(* Schneider Machine Expert - Basic project mojokerto-rev7, file version 2.9.0.0 *)
(* ProjectInformations: Name=New project *)

HARDWARE
  Cpu 0: TM221CE24R
  EthernetConfiguration: NetworkName=M221, IpAllocationMode=FixedAddress, IpAddress=192.168.1.113, SubnetMask=255.255.255.0
  SerialLineConfiguration: Baud=Baud19200, Parity=ParityNone, DataBits=DataBits8, StopBits=StopBits1, PhysicalMedium=PhysicalMediumRs485, TransmissionMode=TransmissionModeIoScannerRtu
  MastTask: UsePeriodScanMode=false, PeriodScan=100
  FastTask: Period=255
  CpuBehavior: StartingMode=StartAsPreviousState, AutoSaveRamOnEeprom=true, WatchdogPeriod=250

SYMBOLS  (address, symbol, comment, settings)
  %M10      VSD1_START  "VSD1 START dari FUXA (pulse)"
  %M11      VSD1_STOP  "VSD1 STOP dari FUXA (pulse)"
  %M12      VSD2_START  "VSD2 START dari FUXA (pulse)"
  %M13      VSD2_STOP  "VSD2 STOP dari FUXA (pulse)"
  %M14      VSD3_START  "VSD3 START dari FUXA (pulse)"
  %M15      VSD3_STOP  "VSD3 STOP dari FUXA (pulse)"
  %M16      VSD4_START  "VSD4 START dari FUXA (pulse)"
  %M17      VSD4_STOP  "VSD4 STOP dari FUXA (pulse)"
  %M18      VSD5_START  "VSD5 START dari FUXA (pulse)"
  %M19      VSD5_STOP  "VSD5 STOP dari FUXA (pulse)"
  %M20      VSD1_RUN_CMD  "VSD1 output RUN aktif"
  %M21      VSD2_RUN_CMD  "VSD2 output RUN aktif"
  %M22      VSD3_RUN_CMD  "VSD3 output RUN aktif"
  %M23      VSD4_RUN_CMD  "VSD4 output RUN aktif"
  %M24      VSD5_RUN_CMD  "VSD5 output RUN aktif"
  %M25      VSD1_RUNNING  "VSD1 berjalan (SW b2)"
  %M26      VSD2_RUNNING  "VSD2 berjalan (SW b2)"
  %M27      VSD3_RUNNING  "VSD3 berjalan (SW b2)"
  %M28      VSD4_RUNNING  "VSD4 berjalan (SW b2)"
  %M29      VSD5_RUNNING  "VSD5 berjalan (SW b2)"
  %M30      MODE_REMOTE  "1 = selector REMOTE (SCADA), 0 = LOCAL (PB panel)"
  %M31      MODE_ESTOP_OK  "Salinan %I0.1 untuk FUXA: 1 = e-stop sehat"
  %M40      VSD1_FAULT  "VSD1 fault (SW b3, comm OK)"
  %M41      VSD2_FAULT  "VSD2 fault (SW b3, comm OK)"
  %M42      VSD3_FAULT  "VSD3 fault (SW b3, comm OK)"
  %M43      VSD4_FAULT  "VSD4 fault (SW b3, comm OK)"
  %M44      VSD5_FAULT  "VSD5 fault (SW b3, comm OK)"
  %M45      VSD1_WARN  "VSD1 warning (SW b7)"
  %M46      VSD2_WARN  "VSD2 warning (SW b7)"
  %M47      VSD3_WARN  "VSD3 warning (SW b7)"
  %M48      VSD4_WARN  "VSD4 warning (SW b7)"
  %M49      VSD5_WARN  "VSD5 warning (SW b7)"
  %M50      VSD1_REMOTE  "VSD1 di REMOTE (SW b9)"
  %M51      VSD2_REMOTE  "VSD2 di REMOTE (SW b9)"
  %M52      VSD3_REMOTE  "VSD3 di REMOTE (SW b9)"
  %M53      VSD4_REMOTE  "VSD4 di REMOTE (SW b9)"
  %M54      VSD5_REMOTE  "VSD5 di REMOTE (SW b9)"
  %M60      VSD1_COMM_OK  "VSD1 IOScanner status = 2"
  %M61      VSD2_COMM_OK  "VSD2 IOScanner status = 2"
  %M62      VSD3_COMM_OK  "VSD3 IOScanner status = 2"
  %M63      VSD4_COMM_OK  "VSD4 IOScanner status = 2"
  %M64      VSD5_COMM_OK  "VSD5 IOScanner status = 2"
  %M65      FLOW_COMM_OK  "Flow meter IOScanner status = 2"
  %M70      VSD1_COMM_LOST  "VSD1 alarm komunikasi putus"
  %M71      VSD2_COMM_LOST  "VSD2 alarm komunikasi putus"
  %M72      VSD3_COMM_LOST  "VSD3 alarm komunikasi putus"
  %M73      VSD4_COMM_LOST  "VSD4 alarm komunikasi putus"
  %M74      VSD5_COMM_LOST  "VSD5 alarm komunikasi putus"
  %M75      FLOW_COMM_LOST  "Flow meter alarm komunikasi putus"
  %M80      FLOW_PIPE_EMPTY  "Flow: pipa kosong"
  %M81      FLOW_COIL_ERR  "Flow: coils excitation error"
  %M82      FLOW_MIN  "Flow: di bawah MIN"
  %M83      FLOW_MAX  "Flow: di atas MAX"
  %M90      VSD3_INSTALLED  "1 = VSD3 sudah terpasang, alarm comm lost VSD3 aktif"
  %M99      WORD_SWAP  "0 = tukar word 32-bit (default), 1 = lurus"
  %M111     RETRY_PULSE  "Pulse auto-retry IOScanner (rev5)"
  %M112     S6_PREV  "%S6 scan sebelumnya (deteksi sisi naik)"
  %S6       SB_TB1S  "Time base of 1 s generated by an internal clock"
  %S13      SB_FIRSTRUN  "Indicates the first controller cycle in RUN mode"
  %S110     SB_IOSCAN1RESET  "Set to 1 to reset the IOScanner on Serial Line 1"
  %SW210    SW_IOSCAN1STATUS  "Contains the IOScanner status of Serial Line 1"
  %MW990    SP_MIN  "Setpoint minimum Hz x10"
  %MW991    SP_MAX  "Setpoint maksimum Hz x10"
  %MW1000   VSD1_SW  "VSD1 status word"
  %MW1001   VSD1_FREQ  "VSD1 frekuensi Hz x10"
  %MW1002   VSD1_CURRENT  "VSD1 arus A x10"
  %MW1003   VSD1_DCBUS  "VSD1 DC bus V"
  %MW1004   VSD1_VOUT  "VSD1 Vout V"
  %MW1005   VSD1_REF_RB  "VSD1 ref1 terbaca Hz x10"
  %MW1006   VSD1_SP  "VSD1 setpoint dari FUXA Hz x10"
  %MW1020   VSD2_SW  "VSD2 status word"
  %MW1021   VSD2_FREQ  "VSD2 frekuensi Hz x10"
  %MW1022   VSD2_CURRENT  "VSD2 arus A x10"
  %MW1023   VSD2_DCBUS  "VSD2 DC bus V"
  %MW1024   VSD2_VOUT  "VSD2 Vout V"
  %MW1025   VSD2_REF_RB  "VSD2 ref1 terbaca Hz x10"
  %MW1026   VSD2_SP  "VSD2 setpoint dari FUXA Hz x10"
  %MW1040   VSD3_SW  "VSD3 status word"
  %MW1041   VSD3_FREQ  "VSD3 frekuensi Hz x10"
  %MW1042   VSD3_CURRENT  "VSD3 arus A x10"
  %MW1043   VSD3_DCBUS  "VSD3 DC bus V"
  %MW1044   VSD3_VOUT  "VSD3 Vout V"
  %MW1045   VSD3_REF_RB  "VSD3 ref1 terbaca Hz x10"
  %MW1046   VSD3_SP  "VSD3 setpoint dari FUXA Hz x10"
  %MW1060   VSD4_SW  "VSD4 status word"
  %MW1061   VSD4_FREQ  "VSD4 frekuensi Hz x10"
  %MW1062   VSD4_CURRENT  "VSD4 arus A x10"
  %MW1063   VSD4_DCBUS  "VSD4 DC bus V"
  %MW1064   VSD4_VOUT  "VSD4 Vout V"
  %MW1065   VSD4_REF_RB  "VSD4 ref1 terbaca Hz x10"
  %MW1066   VSD4_SP  "VSD4 setpoint dari FUXA Hz x10"
  %MW1080   VSD5_SW  "VSD5 status word"
  %MW1081   VSD5_FREQ  "VSD5 frekuensi Hz x10"
  %MW1082   VSD5_CURRENT  "VSD5 arus A x10"
  %MW1083   VSD5_DCBUS  "VSD5 DC bus V"
  %MW1084   VSD5_VOUT  "VSD5 Vout V"
  %MW1085   VSD5_REF_RB  "VSD5 ref1 terbaca Hz x10"
  %MW1086   VSD5_SP  "VSD5 setpoint dari FUXA Hz x10"
  %MW1112   FLOW_TP_INFO  "T+ MSB overflow LSB desimal"
  %MW1113   FLOW_TN_INFO  "T- info"
  %MW1114   FLOW_FLAGS12  "Flag 1/2 reg 0020"
  %MW1115   FLOW_ALARMS  "Jumlah alarm"
  %MW1116   FLOW_BATT  "Baterai %"
  %MW1117   FLOW_FLAGS34  "Flag 3/4 reg 0051"
  %MW1600   VSD1_IOS_STAT  "VSD1 status device IOScanner"
  %MW1601   VSD2_IOS_STAT  "VSD2 status device IOScanner"
  %MW1602   VSD3_IOS_STAT  "VSD3 status device IOScanner"
  %MW1603   FLOW_IOS_STAT  "Flow status device IOScanner"
  %MW1604   VSD4_IOS_STAT  "VSD4 status device IOScanner"
  %MW1605   VSD5_IOS_STAT  "VSD5 status device IOScanner"
  %MW1606   IOS_SL1_STATE  "%SW210: 0 stop 1 init 2 OK 3 sebagian 4 suspend"
  %MW1610   RETRY_SEC_CNT  "Hitungan detik auto-retry IOScanner"
  %MW1611   IOS_RESET_COUNT  "Jumlah reset IOScanner SL1 oleh program"
  %I0.0     SEL_REMOTE  "Selector panel: 1 = REMOTE (start/stop SCADA), 0 = LOCAL (PB panel)"
  %I0.1     ESTOP_OK  "E-stop, kontak NC: 1 = sehat"
  %I0.2     VSD1_PB_ON  "PB ON VSD1 di panel (NO), aktif di LOCAL"
  %I0.3     VSD1_PB_OFF  "PB OFF VSD1 di panel (NC), aktif di LOCAL dan REMOTE, 0 = stop"
  %I0.4     VSD2_PB_ON  "PB ON VSD2 di panel (NO), aktif di LOCAL"
  %I0.5     VSD2_PB_OFF  "PB OFF VSD2 di panel (NC), aktif di LOCAL dan REMOTE, 0 = stop"
  %I0.6     VSD3_PB_ON  "PB ON VSD3 di panel (NO), aktif di LOCAL"
  %I0.7     VSD3_PB_OFF  "PB OFF VSD3 di panel (NC), aktif di LOCAL dan REMOTE, 0 = stop"
  %I0.8     VSD4_PB_ON  "PB ON VSD4 di panel (NO), aktif di LOCAL"
  %I0.9     VSD4_PB_OFF  "PB OFF VSD4 di panel (NC), aktif di LOCAL dan REMOTE, 0 = stop"
  %I0.10    VSD5_PB_ON  "PB ON VSD5 di panel (NO), aktif di LOCAL"
  %I0.11    VSD5_PB_OFF  "PB OFF VSD5 di panel (NC), aktif di LOCAL dan REMOTE, 0 = stop"
  %Q0.0     VSD1_RUN  "Ke DI start VSD1 (ACS550), hardwired"
  %Q0.1     VSD2_RUN  "Ke DI start VSD2 (ACS580), hardwired"
  %Q0.2     VSD3_RUN  "Ke DI start VSD3 (ACS580), hardwired"
  %Q0.3     VSD4_RUN  "Ke DI start VSD4 (ACS580), hardwired"
  %Q0.4     VSD5_RUN  "Ke DI start VSD5 (ACS580), hardwired"
  %IWN100.0.0   [Channel=SW_REF_ACT]
  %IWN100.0.1   [Channel=SW_REF_ACT]
  %IWN100.0.2   [Channel=SW_REF_ACT]
  %IWN100.0.3   [Channel=SW_REF_ACT]
  %IWN100.1.0   [Channel=PAR_0103_0111]
  %IWN100.1.1   [Channel=PAR_0103_0111]
  %IWN100.1.2   [Channel=PAR_0103_0111]
  %IWN100.1.3   [Channel=PAR_0103_0111]
  %IWN100.1.4   [Channel=PAR_0103_0111]
  %IWN100.1.5   [Channel=PAR_0103_0111]
  %IWN100.1.6   [Channel=PAR_0103_0111]
  %IWN100.1.7   [Channel=PAR_0103_0111]
  %IWN100.1.8   [Channel=PAR_0103_0111]
  %IWN101.0.0   [Channel=SW_REF_ACT]
  %IWN101.0.1   [Channel=SW_REF_ACT]
  %IWN101.0.2   [Channel=SW_REF_ACT]
  %IWN101.0.3   [Channel=SW_REF_ACT]
  %IWN101.1.0   [Channel=CURRENT_32]
  %IWN101.1.1   [Channel=CURRENT_32]
  %IWN101.2.0   [Channel=DC_BUS]
  %IWN101.3.0   [Channel=VOUT]
  %IWN102.0.0   [Channel=SW_REF_ACT]
  %IWN102.0.1   [Channel=SW_REF_ACT]
  %IWN102.0.2   [Channel=SW_REF_ACT]
  %IWN102.0.3   [Channel=SW_REF_ACT]
  %IWN102.1.0   [Channel=CURRENT_32]
  %IWN102.1.1   [Channel=CURRENT_32]
  %IWN102.2.0   [Channel=DC_BUS]
  %IWN102.3.0   [Channel=VOUT]
  %IWN103.0.0   [Channel=FLOW_TOT_FLAGS]
  %IWN103.0.1   [Channel=FLOW_TOT_FLAGS]
  %IWN103.0.2   [Channel=FLOW_TOT_FLAGS]
  %IWN103.0.3   [Channel=FLOW_TOT_FLAGS]
  %IWN103.0.4   [Channel=FLOW_TOT_FLAGS]
  %IWN103.0.5   [Channel=FLOW_TOT_FLAGS]
  %IWN103.0.6   [Channel=FLOW_TOT_FLAGS]
  %IWN103.0.7   [Channel=FLOW_TOT_FLAGS]
  %IWN103.0.8   [Channel=FLOW_TOT_FLAGS]
  %IWN103.0.9   [Channel=FLOW_TOT_FLAGS]
  %IWN103.0.10   [Channel=FLOW_TOT_FLAGS]
  %IWN103.0.11   [Channel=FLOW_TOT_FLAGS]
  %IWN103.0.12   [Channel=FLOW_TOT_FLAGS]
  %IWN103.0.13   [Channel=FLOW_TOT_FLAGS]
  %IWN103.0.14   [Channel=FLOW_TOT_FLAGS]
  %IWN103.0.15   [Channel=FLOW_TOT_FLAGS]
  %IWN103.0.16   [Channel=FLOW_TOT_FLAGS]
  %IWN103.0.17   [Channel=FLOW_TOT_FLAGS]
  %IWN103.0.18   [Channel=FLOW_TOT_FLAGS]
  %IWN103.1.0   [Channel=BATT_ALM_LPS]
  %IWN103.1.1   [Channel=BATT_ALM_LPS]
  %IWN103.1.2   [Channel=BATT_ALM_LPS]
  %IWN103.1.3   [Channel=BATT_ALM_LPS]
  %IWN103.1.4   [Channel=BATT_ALM_LPS]
  %IWN103.1.5   [Channel=BATT_ALM_LPS]
  %IWN103.1.6   [Channel=BATT_ALM_LPS]
  %IWN103.1.7   [Channel=BATT_ALM_LPS]
  %IWN103.1.8   [Channel=BATT_ALM_LPS]
  %IWN103.1.9   [Channel=BATT_ALM_LPS]
  %IWN103.2.0   [Channel=FLAGS_3_4]
  %IWN104.0.0   [Channel=SW_REF_ACT]
  %IWN104.0.1   [Channel=SW_REF_ACT]
  %IWN104.0.2   [Channel=SW_REF_ACT]
  %IWN104.0.3   [Channel=SW_REF_ACT]
  %IWN104.1.0   [Channel=CURRENT_32]
  %IWN104.1.1   [Channel=CURRENT_32]
  %IWN104.2.0   [Channel=DC_BUS]
  %IWN104.3.0   [Channel=VOUT]
  %IWN105.0.0   [Channel=SW_REF_ACT]
  %IWN105.0.1   [Channel=SW_REF_ACT]
  %IWN105.0.2   [Channel=SW_REF_ACT]
  %IWN105.0.3   [Channel=SW_REF_ACT]
  %IWN105.1.0   [Channel=CURRENT_32]
  %IWN105.1.1   [Channel=CURRENT_32]
  %IWN105.2.0   [Channel=DC_BUS]
  %IWN105.3.0   [Channel=VOUT]
  %QWN100.2.0   [Channel=REF1_WRITE]
  %QWN101.4.0   [Channel=REF1_WRITE]
  %QWN102.4.0   [Channel=REF1_WRITE]
  %QWN104.4.0   [Channel=REF1_WRITE]
  %QWN105.4.0   [Channel=REF1_WRITE]

POU Mojokerto
  (* SectionNumber=0 *)

// Rung 0: INIT
// Cold start: batas setpoint default 0..50,0 Hz (x10)
  LD %S13                 (* SB_FIRSTRUN - Siklus pertama setelah start *)
  [ %MW990 := 0 ]         (* SP_MIN - SP_MIN Hz x10 *)
  [ %MW991 := 500 ]       (* SP_MAX - SP_MAX Hz x10 *)
  // as ST:
  //   IF SB_FIRSTRUN THEN SP_MIN := 0; END_IF;
  //   IF SB_FIRSTRUN THEN SP_MAX := 500; END_IF;

// Rung 1: RAW_VSD1
// Salin data IOScanner VSD1 (ACS550, slave ID 1) ke %MW1300
  LD 1                    (* Selalu *)
  [ %MW1300 := %IWN100.0.0 ](* ref1 *)
  [ %MW1301 := %IWN100.0.1 ](* ref2 *)
  [ %MW1302 := %IWN100.0.2 ](* status word *)
  [ %MW1303 := %IWN100.0.3 ](* act1 *)
  [ %MW1304 := %IWN100.1.0 ](* par 0103 *)
  [ %MW1305 := %IWN100.1.1 ](* par 0104 *)
  [ %MW1306 := %IWN100.1.2 ](* par 0105 *)
  [ %MW1307 := %IWN100.1.3 ](* par 0106 *)
  [ %MW1308 := %IWN100.1.4 ](* par 0107 *)
  [ %MW1309 := %IWN100.1.5 ](* par 0108 *)
  [ %MW1310 := %IWN100.1.6 ](* par 0109 *)
  [ %MW1311 := %IWN100.1.7 ](* par 0110 *)
  [ %MW1312 := %IWN100.1.8 ](* par 0111 *)
  [ %MW1600 := %IWNS100 ] (* VSD1_IOS_STAT - status device IOScanner (2 = OK) *)
  // as ST:
  //   %MW1300 := %IWN100.0.0;
  //   %MW1301 := %IWN100.0.1;
  //   %MW1302 := %IWN100.0.2;
  //   %MW1303 := %IWN100.0.3;
  //   %MW1304 := %IWN100.1.0;
  //   %MW1305 := %IWN100.1.1;
  //   %MW1306 := %IWN100.1.2;
  //   %MW1307 := %IWN100.1.3;
  //   %MW1308 := %IWN100.1.4;
  //   %MW1309 := %IWN100.1.5;
  //   %MW1310 := %IWN100.1.6;
  //   %MW1311 := %IWN100.1.7;
  //   %MW1312 := %IWN100.1.8;
  //   VSD1_IOS_STAT := %IWNS100;

// Rung 2: RAW_VSD2
// Salin data IOScanner VSD2 (ACS580, slave ID 2) ke %MW1340
  LD 1                    (* Selalu *)
  [ %MW1340 := %IWN101.0.0 ](* ref1 *)
  [ %MW1341 := %IWN101.0.1 ](* ref2 *)
  [ %MW1342 := %IWN101.0.2 ](* status word *)
  [ %MW1343 := %IWN101.0.3 ](* act1 *)
  [ %MW1344 := %IWN101.1.0 ](* 01.07 arus word 1 *)
  [ %MW1345 := %IWN101.1.1 ](* 01.07 arus word 2 *)
  [ %MW1346 := %IWN101.2.0 ](* 01.11 DC bus *)
  [ %MW1347 := %IWN101.3.0 ](* 01.13 Vout *)
  [ %MW1601 := %IWNS101 ] (* VSD2_IOS_STAT - status device IOScanner (2 = OK) *)
  // as ST:
  //   %MW1340 := %IWN101.0.0;
  //   %MW1341 := %IWN101.0.1;
  //   %MW1342 := %IWN101.0.2;
  //   %MW1343 := %IWN101.0.3;
  //   %MW1344 := %IWN101.1.0;
  //   %MW1345 := %IWN101.1.1;
  //   %MW1346 := %IWN101.2.0;
  //   %MW1347 := %IWN101.3.0;
  //   VSD2_IOS_STAT := %IWNS101;

// Rung 3: RAW_VSD3
// Salin data IOScanner VSD3 (ACS580, slave ID 3) ke %MW1380
  LD 1                    (* Selalu *)
  [ %MW1380 := %IWN102.0.0 ](* ref1 *)
  [ %MW1381 := %IWN102.0.1 ](* ref2 *)
  [ %MW1382 := %IWN102.0.2 ](* status word *)
  [ %MW1383 := %IWN102.0.3 ](* act1 *)
  [ %MW1384 := %IWN102.1.0 ](* 01.07 arus word 1 *)
  [ %MW1385 := %IWN102.1.1 ](* 01.07 arus word 2 *)
  [ %MW1386 := %IWN102.2.0 ](* 01.11 DC bus *)
  [ %MW1387 := %IWN102.3.0 ](* 01.13 Vout *)
  [ %MW1602 := %IWNS102 ] (* VSD3_IOS_STAT - status device IOScanner (2 = OK) *)
  // as ST:
  //   %MW1380 := %IWN102.0.0;
  //   %MW1381 := %IWN102.0.1;
  //   %MW1382 := %IWN102.0.2;
  //   %MW1383 := %IWN102.0.3;
  //   %MW1384 := %IWN102.1.0;
  //   %MW1385 := %IWN102.1.1;
  //   %MW1386 := %IWN102.2.0;
  //   %MW1387 := %IWN102.3.0;
  //   VSD3_IOS_STAT := %IWNS102;

// Rung 4: RAW_VSD4
// Salin data IOScanner VSD4 (ACS580, slave ID 5) ke %MW1460
  LD 1                    (* Selalu *)
  [ %MW1460 := %IWN104.0.0 ](* ref1 *)
  [ %MW1461 := %IWN104.0.1 ](* ref2 *)
  [ %MW1462 := %IWN104.0.2 ](* status word *)
  [ %MW1463 := %IWN104.0.3 ](* act1 *)
  [ %MW1464 := %IWN104.1.0 ](* 01.07 arus word 1 *)
  [ %MW1465 := %IWN104.1.1 ](* 01.07 arus word 2 *)
  [ %MW1466 := %IWN104.2.0 ](* 01.11 DC bus *)
  [ %MW1467 := %IWN104.3.0 ](* 01.13 Vout *)
  [ %MW1604 := %IWNS104 ] (* VSD4_IOS_STAT - status device IOScanner (2 = OK) *)
  // as ST:
  //   %MW1460 := %IWN104.0.0;
  //   %MW1461 := %IWN104.0.1;
  //   %MW1462 := %IWN104.0.2;
  //   %MW1463 := %IWN104.0.3;
  //   %MW1464 := %IWN104.1.0;
  //   %MW1465 := %IWN104.1.1;
  //   %MW1466 := %IWN104.2.0;
  //   %MW1467 := %IWN104.3.0;
  //   VSD4_IOS_STAT := %IWNS104;

// Rung 5: RAW_VSD5
// Salin data IOScanner VSD5 (ACS580, slave ID 6) ke %MW1500
  LD 1                    (* Selalu *)
  [ %MW1500 := %IWN105.0.0 ](* ref1 *)
  [ %MW1501 := %IWN105.0.1 ](* ref2 *)
  [ %MW1502 := %IWN105.0.2 ](* status word *)
  [ %MW1503 := %IWN105.0.3 ](* act1 *)
  [ %MW1504 := %IWN105.1.0 ](* 01.07 arus word 1 *)
  [ %MW1505 := %IWN105.1.1 ](* 01.07 arus word 2 *)
  [ %MW1506 := %IWN105.2.0 ](* 01.11 DC bus *)
  [ %MW1507 := %IWN105.3.0 ](* 01.13 Vout *)
  [ %MW1605 := %IWNS105 ] (* VSD5_IOS_STAT - status device IOScanner (2 = OK) *)
  // as ST:
  //   %MW1500 := %IWN105.0.0;
  //   %MW1501 := %IWN105.0.1;
  //   %MW1502 := %IWN105.0.2;
  //   %MW1503 := %IWN105.0.3;
  //   %MW1504 := %IWN105.1.0;
  //   %MW1505 := %IWN105.1.1;
  //   %MW1506 := %IWN105.2.0;
  //   %MW1507 := %IWN105.3.0;
  //   VSD5_IOS_STAT := %IWNS105;

// Rung 6: RAW_FLOW
// Salin data IOScanner flow meter MV145 (slave ID 4) ke %MW1420
  LD 1                    (* Selalu *)
  [ %MW1420 := %IWN103.0.0 ](* MV145 reg 0002 *)
  [ %MW1421 := %IWN103.0.1 ](* MV145 reg 0003 *)
  [ %MW1422 := %IWN103.0.2 ](* MV145 reg 0004 *)
  [ %MW1423 := %IWN103.0.3 ](* MV145 reg 0005 *)
  [ %MW1424 := %IWN103.0.4 ](* MV145 reg 0006 *)
  [ %MW1425 := %IWN103.0.5 ](* MV145 reg 0007 *)
  [ %MW1426 := %IWN103.0.6 ](* MV145 reg 0008 *)
  [ %MW1427 := %IWN103.0.7 ](* MV145 reg 0009 *)
  [ %MW1428 := %IWN103.0.8 ](* MV145 reg 0010 *)
  [ %MW1429 := %IWN103.0.9 ](* MV145 reg 0011 *)
  [ %MW1430 := %IWN103.0.10 ](* MV145 reg 0012 *)
  [ %MW1431 := %IWN103.0.11 ](* MV145 reg 0013 *)
  [ %MW1432 := %IWN103.0.12 ](* MV145 reg 0014 *)
  [ %MW1433 := %IWN103.0.13 ](* MV145 reg 0015 *)
  [ %MW1434 := %IWN103.0.14 ](* MV145 reg 0016 *)
  [ %MW1435 := %IWN103.0.15 ](* MV145 reg 0017 *)
  [ %MW1436 := %IWN103.0.16 ](* MV145 reg 0018 *)
  [ %MW1437 := %IWN103.0.17 ](* MV145 reg 0019 *)
  [ %MW1438 := %IWN103.0.18 ](* MV145 reg 0020 *)
  [ %MW1440 := %IWN103.1.0 ](* MV145 reg 0027 *)
  [ %MW1441 := %IWN103.1.1 ](* MV145 reg 0028 *)
  [ %MW1442 := %IWN103.1.2 ](* MV145 reg 0029 *)
  [ %MW1443 := %IWN103.1.3 ](* MV145 reg 0030 *)
  [ %MW1444 := %IWN103.1.4 ](* MV145 reg 0031 *)
  [ %MW1445 := %IWN103.1.5 ](* MV145 reg 0032 *)
  [ %MW1446 := %IWN103.1.6 ](* MV145 reg 0033 *)
  [ %MW1447 := %IWN103.1.7 ](* MV145 reg 0034 *)
  [ %MW1448 := %IWN103.1.8 ](* MV145 reg 0035 *)
  [ %MW1449 := %IWN103.1.9 ](* MV145 reg 0036 *)
  [ %MW1450 := %IWN103.2.0 ](* MV145 reg 0051 *)
  [ %MW1603 := %IWNS103 ] (* FLOW_IOS_STAT - status device IOScanner flow (2 = OK) *)
  // as ST:
  //   %MW1420 := %IWN103.0.0;
  //   %MW1421 := %IWN103.0.1;
  //   %MW1422 := %IWN103.0.2;
  //   %MW1423 := %IWN103.0.3;
  //   %MW1424 := %IWN103.0.4;
  //   %MW1425 := %IWN103.0.5;
  //   %MW1426 := %IWN103.0.6;
  //   %MW1427 := %IWN103.0.7;
  //   %MW1428 := %IWN103.0.8;
  //   %MW1429 := %IWN103.0.9;
  //   %MW1430 := %IWN103.0.10;
  //   %MW1431 := %IWN103.0.11;
  //   %MW1432 := %IWN103.0.12;
  //   %MW1433 := %IWN103.0.13;
  //   %MW1434 := %IWN103.0.14;
  //   %MW1435 := %IWN103.0.15;
  //   %MW1436 := %IWN103.0.16;
  //   %MW1437 := %IWN103.0.17;
  //   %MW1438 := %IWN103.0.18;
  //   %MW1440 := %IWN103.1.0;
  //   %MW1441 := %IWN103.1.1;
  //   %MW1442 := %IWN103.1.2;
  //   %MW1443 := %IWN103.1.3;
  //   %MW1444 := %IWN103.1.4;
  //   %MW1445 := %IWN103.1.5;
  //   %MW1446 := %IWN103.1.6;
  //   %MW1447 := %IWN103.1.7;
  //   %MW1448 := %IWN103.1.8;
  //   %MW1449 := %IWN103.1.9;
  //   %MW1450 := %IWN103.2.0;
  //   FLOW_IOS_STAT := %IWNS103;

// Rung 7: COMM_OK_SET_VSD1
// VSD1: komunikasi OK saat status device IOScanner = 2
  LD [ %MW1600 = 2 ]      (* VSD1_IOS_STAT *)
  S %M60                  (* VSD1_COMM_OK *)
  // as ST:
  //   IF VSD1_IOS_STAT = 2 THEN VSD1_COMM_OK := TRUE; END_IF;

// Rung 8: COMM_OK_RST_VSD1
// VSD1: komunikasi putus saat status bukan 2 dan bukan 1 (1 = init sesudah reset, abaikan)
  LD [ %MW1600 <> 2 ]     (* VSD1_IOS_STAT *)
  AND [ %MW1600 <> 1 ]    (* VSD1_IOS_STAT *)
  R %M60                  (* VSD1_COMM_OK *)
  // as ST:
  //   IF VSD1_IOS_STAT <> 2 AND VSD1_IOS_STAT <> 1 THEN VSD1_COMM_OK := FALSE; END_IF;

// Rung 9: COMM_OK_SET_VSD2
// VSD2: komunikasi OK saat status device IOScanner = 2
  LD [ %MW1601 = 2 ]      (* VSD2_IOS_STAT *)
  S %M61                  (* VSD2_COMM_OK *)
  // as ST:
  //   IF VSD2_IOS_STAT = 2 THEN VSD2_COMM_OK := TRUE; END_IF;

// Rung 10: COMM_OK_RST_VSD2
// VSD2: komunikasi putus saat status bukan 2 dan bukan 1 (1 = init sesudah reset, abaikan)
  LD [ %MW1601 <> 2 ]     (* VSD2_IOS_STAT *)
  AND [ %MW1601 <> 1 ]    (* VSD2_IOS_STAT *)
  R %M61                  (* VSD2_COMM_OK *)
  // as ST:
  //   IF VSD2_IOS_STAT <> 2 AND VSD2_IOS_STAT <> 1 THEN VSD2_COMM_OK := FALSE; END_IF;

// Rung 11: COMM_OK_SET_VSD3
// VSD3: komunikasi OK saat status device IOScanner = 2
  LD [ %MW1602 = 2 ]      (* VSD3_IOS_STAT *)
  S %M62                  (* VSD3_COMM_OK *)
  // as ST:
  //   IF VSD3_IOS_STAT = 2 THEN VSD3_COMM_OK := TRUE; END_IF;

// Rung 12: COMM_OK_RST_VSD3
// VSD3: komunikasi putus saat status bukan 2 dan bukan 1 (1 = init sesudah reset, abaikan)
  LD [ %MW1602 <> 2 ]     (* VSD3_IOS_STAT *)
  AND [ %MW1602 <> 1 ]    (* VSD3_IOS_STAT *)
  R %M62                  (* VSD3_COMM_OK *)
  // as ST:
  //   IF VSD3_IOS_STAT <> 2 AND VSD3_IOS_STAT <> 1 THEN VSD3_COMM_OK := FALSE; END_IF;

// Rung 13: COMM_OK_SET_FLOW
// FLOW: komunikasi OK saat status device IOScanner = 2
  LD [ %MW1603 = 2 ]      (* FLOW_IOS_STAT *)
  S %M65                  (* FLOW_COMM_OK *)
  // as ST:
  //   IF FLOW_IOS_STAT = 2 THEN FLOW_COMM_OK := TRUE; END_IF;

// Rung 14: COMM_OK_RST_FLOW
// FLOW: komunikasi putus saat status bukan 2 dan bukan 1 (1 = init sesudah reset, abaikan)
  LD [ %MW1603 <> 2 ]     (* FLOW_IOS_STAT *)
  AND [ %MW1603 <> 1 ]    (* FLOW_IOS_STAT *)
  R %M65                  (* FLOW_COMM_OK *)
  // as ST:
  //   IF FLOW_IOS_STAT <> 2 AND FLOW_IOS_STAT <> 1 THEN FLOW_COMM_OK := FALSE; END_IF;

// Rung 15: COMM_OK_SET_VSD4
// VSD4: komunikasi OK saat status device IOScanner = 2
  LD [ %MW1604 = 2 ]      (* VSD4_IOS_STAT *)
  S %M63                  (* VSD4_COMM_OK *)
  // as ST:
  //   IF VSD4_IOS_STAT = 2 THEN VSD4_COMM_OK := TRUE; END_IF;

// Rung 16: COMM_OK_RST_VSD4
// VSD4: komunikasi putus saat status bukan 2 dan bukan 1 (1 = init sesudah reset, abaikan)
  LD [ %MW1604 <> 2 ]     (* VSD4_IOS_STAT *)
  AND [ %MW1604 <> 1 ]    (* VSD4_IOS_STAT *)
  R %M63                  (* VSD4_COMM_OK *)
  // as ST:
  //   IF VSD4_IOS_STAT <> 2 AND VSD4_IOS_STAT <> 1 THEN VSD4_COMM_OK := FALSE; END_IF;

// Rung 17: COMM_OK_SET_VSD5
// VSD5: komunikasi OK saat status device IOScanner = 2
  LD [ %MW1605 = 2 ]      (* VSD5_IOS_STAT *)
  S %M64                  (* VSD5_COMM_OK *)
  // as ST:
  //   IF VSD5_IOS_STAT = 2 THEN VSD5_COMM_OK := TRUE; END_IF;

// Rung 18: COMM_OK_RST_VSD5
// VSD5: komunikasi putus saat status bukan 2 dan bukan 1 (1 = init sesudah reset, abaikan)
  LD [ %MW1605 <> 2 ]     (* VSD5_IOS_STAT *)
  AND [ %MW1605 <> 1 ]    (* VSD5_IOS_STAT *)
  R %M64                  (* VSD5_COMM_OK *)
  // as ST:
  //   IF VSD5_IOS_STAT <> 2 AND VSD5_IOS_STAT <> 1 THEN VSD5_COMM_OK := FALSE; END_IF;

// Rung 19: IOS_STATE
// Salin %SW210 (status IOScanner SL1: 0 stop, 1 init, 2 operasional, 3 sebagian, 4 suspend) untuk FUXA/diagnosa
  LD 1
  [ %MW1606 := %SW210 ]   (* IOS_SL1_STATE, SW_IOSCAN1STATUS *)
  // as ST:
  //   IOS_SL1_STATE := SW_IOSCAN1STATUS;

// Rung 20: RETRY_SEC
// Hitung detik: %S6 (basis waktu 1 s) = 1 dan scan sebelumnya 0 (%M112)
  LD %S6                  (* SB_TB1S *)
  ANDN %M112              (* S6_PREV - %S6 scan sebelumnya *)
  [ %MW1610 := %MW1610 + 1 ](* RETRY_SEC_CNT, RETRY_SEC_CNT *)
  // as ST:
  //   IF SB_TB1S AND NOT S6_PREV THEN RETRY_SEC_CNT := RETRY_SEC_CNT + 1; END_IF;

// Rung 21: RETRY_SEC_MEM
// Simpan %S6 untuk deteksi sisi naik di scan berikutnya
  LD %S6                  (* SB_TB1S *)
  ST %M112                (* S6_PREV *)
  // as ST:
  //   S6_PREV := SB_TB1S;

// Rung 22: RETRY_PULSE
// Pulse satu scan tiap 15 detik
  LD [ %MW1610 >= 15 ]    (* RETRY_SEC_CNT *)
  ST %M111                (* RETRY_PULSE *)
  // as ST:
  //   RETRY_PULSE := RETRY_SEC_CNT >= 15;

// Rung 23: RETRY_CNT_CLR
// Nol-kan hitungan detik setelah pulse
  LD %M111                (* RETRY_PULSE *)
  [ %MW1610 := 0 ]        (* RETRY_SEC_CNT *)
  // as ST:
  //   IF RETRY_PULSE THEN RETRY_SEC_CNT := 0; END_IF;

// Rung 24: RETRY_RESET
// IOScanner tidak operasional penuh -> reset IOScanner SL1 (%S110) + hitung jumlah reset
  LD %M111                (* RETRY_PULSE *)
  AND [ %SW210 <> 2 ]     (* SW_IOSCAN1STATUS *)
  S %S110                 (* SB_IOSCAN1RESET - reset Modbus Serial IOScanner SL1 *)
  [ %MW1611 := %MW1611 + 1 ](* IOS_RESET_COUNT, IOS_RESET_COUNT - jumlah reset (diagnosa) *)
  // as ST:
  //   IF RETRY_PULSE AND SW_IOSCAN1STATUS <> 2 THEN SB_IOSCAN1RESET := TRUE; END_IF;
  //   IF RETRY_PULSE AND SW_IOSCAN1STATUS <> 2 THEN IOS_RESET_COUNT := IOS_RESET_COUNT + 1; END_IF;

// Rung 25: RETRY_RESET_CLR
// Pengaman: kalau sistem belum menurunkan %S110 setelah 3 s, turunkan
  LD %S110                (* SB_IOSCAN1RESET *)
  AND [ %MW1610 >= 3 ]    (* RETRY_SEC_CNT *)
  R %S110                 (* SB_IOSCAN1RESET *)
  // as ST:
  //   IF SB_IOSCAN1RESET AND RETRY_SEC_CNT >= 3 THEN SB_IOSCAN1RESET := FALSE; END_IF;

// Rung 26: COMM_LOST
// Alarm komunikasi putus (FUXA). VSD3 hanya bila %M90 = 1 (drive sudah terpasang)
  LDN %M60                (* VSD1_COMM_OK *)
  ST %M70                 (* VSD1_COMM_LOST - VSD1 comm lost *)
  // as ST:
  //   VSD1_COMM_LOST := NOT VSD1_COMM_OK;

// Rung 27: COMM_LOST_VSD2
  LDN %M61                (* VSD2_COMM_OK *)
  ST %M71                 (* VSD2_COMM_LOST *)
  // as ST:
  //   VSD2_COMM_LOST := NOT VSD2_COMM_OK;

// Rung 28: COMM_LOST_VSD3
// VSD3 belum terpasang: alarm hanya aktif kalau %M90 = 1
  LD %M90                 (* VSD3_INSTALLED - VSD3 terpasang *)
  ANDN %M62               (* VSD3_COMM_OK *)
  ST %M72                 (* VSD3_COMM_LOST *)
  // as ST:
  //   VSD3_COMM_LOST := VSD3_INSTALLED AND NOT VSD3_COMM_OK;

// Rung 29: COMM_LOST_VSD4
  LDN %M63                (* VSD4_COMM_OK *)
  ST %M73                 (* VSD4_COMM_LOST *)
  // as ST:
  //   VSD4_COMM_LOST := NOT VSD4_COMM_OK;

// Rung 30: COMM_LOST_VSD5
  LDN %M64                (* VSD5_COMM_OK *)
  ST %M74                 (* VSD5_COMM_LOST *)
  // as ST:
  //   VSD5_COMM_LOST := NOT VSD5_COMM_OK;

// Rung 31: COMM_LOST_FLOW
  LDN %M65                (* FLOW_COMM_OK *)
  ST %M75                 (* FLOW_COMM_LOST *)
  // as ST:
  //   FLOW_COMM_LOST := NOT FLOW_COMM_OK;

// Rung 32: WORD32_SWAP
// Rakit float/32-bit flow meter + arus ACS580, word ditukar. Uji saat commissioning: %MF1100 harus = flow di layar MV145
  LDN %M99                (* WORD_SWAP - WORD_SWAP = 0 -> tukar word *)
  [ %MW1100 := %MW1423 ]
  [ %MW1101 := %MW1422 ]
  [ %MW1102 := %MW1449 ]
  [ %MW1103 := %MW1448 ]
  [ %MW1104 := %MW1421 ]
  [ %MW1105 := %MW1420 ]
  [ %MW1106 := %MW1425 ]
  [ %MW1107 := %MW1424 ]
  [ %MW1108 := %MW1427 ]
  [ %MW1109 := %MW1426 ]
  [ %MW1110 := %MW1433 ]
  [ %MW1111 := %MW1432 ]
  [ %MW1210 := %MW1345 ]
  [ %MW1211 := %MW1344 ]
  [ %MW1212 := %MW1385 ]
  [ %MW1213 := %MW1384 ]
  [ %MW1214 := %MW1465 ]
  [ %MW1215 := %MW1464 ]
  [ %MW1216 := %MW1505 ]
  [ %MW1217 := %MW1504 ]
  // as ST:
  //   IF NOT WORD_SWAP THEN %MW1100 := %MW1423; END_IF;
  //   IF NOT WORD_SWAP THEN %MW1101 := %MW1422; END_IF;
  //   IF NOT WORD_SWAP THEN %MW1102 := %MW1449; END_IF;
  //   IF NOT WORD_SWAP THEN %MW1103 := %MW1448; END_IF;
  //   IF NOT WORD_SWAP THEN %MW1104 := %MW1421; END_IF;
  //   IF NOT WORD_SWAP THEN %MW1105 := %MW1420; END_IF;
  //   IF NOT WORD_SWAP THEN %MW1106 := %MW1425; END_IF;
  //   IF NOT WORD_SWAP THEN %MW1107 := %MW1424; END_IF;
  //   IF NOT WORD_SWAP THEN %MW1108 := %MW1427; END_IF;
  //   IF NOT WORD_SWAP THEN %MW1109 := %MW1426; END_IF;
  //   IF NOT WORD_SWAP THEN %MW1110 := %MW1433; END_IF;
  //   IF NOT WORD_SWAP THEN %MW1111 := %MW1432; END_IF;
  //   IF NOT WORD_SWAP THEN %MW1210 := %MW1345; END_IF;
  //   IF NOT WORD_SWAP THEN %MW1211 := %MW1344; END_IF;
  //   IF NOT WORD_SWAP THEN %MW1212 := %MW1385; END_IF;
  //   IF NOT WORD_SWAP THEN %MW1213 := %MW1384; END_IF;
  //   IF NOT WORD_SWAP THEN %MW1214 := %MW1465; END_IF;
  //   IF NOT WORD_SWAP THEN %MW1215 := %MW1464; END_IF;
  //   IF NOT WORD_SWAP THEN %MW1216 := %MW1505; END_IF;
  //   IF NOT WORD_SWAP THEN %MW1217 := %MW1504; END_IF;

// Rung 33: WORD32_STRAIGHT
// Sama, tanpa tukar word (pakai kalau %M99 = 1)
  LD %M99                 (* WORD_SWAP - WORD_SWAP = 1 -> tanpa tukar *)
  [ %MW1100 := %MW1422 ]
  [ %MW1101 := %MW1423 ]
  [ %MW1102 := %MW1448 ]
  [ %MW1103 := %MW1449 ]
  [ %MW1104 := %MW1420 ]
  [ %MW1105 := %MW1421 ]
  [ %MW1106 := %MW1424 ]
  [ %MW1107 := %MW1425 ]
  [ %MW1108 := %MW1426 ]
  [ %MW1109 := %MW1427 ]
  [ %MW1110 := %MW1432 ]
  [ %MW1111 := %MW1433 ]
  [ %MW1210 := %MW1344 ]
  [ %MW1211 := %MW1345 ]
  [ %MW1212 := %MW1384 ]
  [ %MW1213 := %MW1385 ]
  [ %MW1214 := %MW1464 ]
  [ %MW1215 := %MW1465 ]
  [ %MW1216 := %MW1504 ]
  [ %MW1217 := %MW1505 ]
  // as ST:
  //   IF WORD_SWAP THEN %MW1100 := %MW1422; END_IF;
  //   IF WORD_SWAP THEN %MW1101 := %MW1423; END_IF;
  //   IF WORD_SWAP THEN %MW1102 := %MW1448; END_IF;
  //   IF WORD_SWAP THEN %MW1103 := %MW1449; END_IF;
  //   IF WORD_SWAP THEN %MW1104 := %MW1420; END_IF;
  //   IF WORD_SWAP THEN %MW1105 := %MW1421; END_IF;
  //   IF WORD_SWAP THEN %MW1106 := %MW1424; END_IF;
  //   IF WORD_SWAP THEN %MW1107 := %MW1425; END_IF;
  //   IF WORD_SWAP THEN %MW1108 := %MW1426; END_IF;
  //   IF WORD_SWAP THEN %MW1109 := %MW1427; END_IF;
  //   IF WORD_SWAP THEN %MW1110 := %MW1432; END_IF;
  //   IF WORD_SWAP THEN %MW1111 := %MW1433; END_IF;
  //   IF WORD_SWAP THEN %MW1210 := %MW1344; END_IF;
  //   IF WORD_SWAP THEN %MW1211 := %MW1345; END_IF;
  //   IF WORD_SWAP THEN %MW1212 := %MW1384; END_IF;
  //   IF WORD_SWAP THEN %MW1213 := %MW1385; END_IF;
  //   IF WORD_SWAP THEN %MW1214 := %MW1464; END_IF;
  //   IF WORD_SWAP THEN %MW1215 := %MW1465; END_IF;
  //   IF WORD_SWAP THEN %MW1216 := %MW1504; END_IF;
  //   IF WORD_SWAP THEN %MW1217 := %MW1505; END_IF;

// Rung 34: FLOW_WORDS
// Flow meter: info totalizer, flag, alarm, baterai
  LD 1
  [ %MW1112 := %MW1428 ]  (* FLOW_TP_INFO - T+ info: MSB overflow, LSB jumlah desimal *)
  [ %MW1113 := %MW1434 ]  (* FLOW_TN_INFO - T- info *)
  [ %MW1114 := %MW1438 ]  (* FLOW_FLAGS12 - flag 1 (MSB) / flag 2 (LSB), reg 0020 *)
  [ %MW1115 := %MW1447 ]  (* FLOW_ALARMS - jumlah alarm aktif, reg 0034 *)
  [ %MW1116 := %MW1440 ]  (* FLOW_BATT - baterai %, reg 0027 *)
  [ %MW1117 := %MW1450 ]  (* FLOW_FLAGS34 - flag 3/4, reg 0051 *)
  // as ST:
  //   FLOW_TP_INFO := %MW1428;
  //   FLOW_TN_INFO := %MW1434;
  //   FLOW_FLAGS12 := %MW1438;
  //   FLOW_ALARMS := %MW1447;
  //   FLOW_BATT := %MW1440;
  //   FLOW_FLAGS34 := %MW1450;

// Rung 35: FLOW_ALM_EMPTY
// Flow: pipa kosong (flag 2 bit 0)
  LD %MW1114:X0           (* FLOW_FLAGS12 *)
  ST %M80                 (* FLOW_PIPE_EMPTY *)
  // as ST:
  //   FLOW_PIPE_EMPTY := FLOW_FLAGS12:X0;

// Rung 36: FLOW_ALM_COIL
// Flow: coils excitation error (flag 2 bit 1)
  LD %MW1114:X1           (* FLOW_FLAGS12 *)
  ST %M81                 (* FLOW_COIL_ERR *)
  // as ST:
  //   FLOW_COIL_ERR := FLOW_FLAGS12:X1;

// Rung 37: FLOW_ALM_MIN
// Flow: di bawah ambang MIN (flag 1 bit 7)
  LD %MW1114:X15          (* FLOW_FLAGS12 *)
  ST %M82                 (* FLOW_MIN *)
  // as ST:
  //   FLOW_MIN := FLOW_FLAGS12:X15;

// Rung 38: FLOW_ALM_MAX
// Flow: di atas ambang MAX (flag 1 bit 6)
  LD %MW1114:X14          (* FLOW_FLAGS12 *)
  ST %M83                 (* FLOW_MAX *)
  // as ST:
  //   FLOW_MAX := FLOW_FLAGS12:X14;

// Rung 39: SCALE_VSD1
// VSD1 ACS550 -> FUXA (sudah 0,1 Hz / 0,1 A dari drive)
  LD 1
  [ %MW1000 := %MW1302 ]  (* VSD1_SW - status word *)
  [ %MW1001 := %MW1304 ]  (* VSD1_FREQ - par 0103 freq Hz x10 *)
  [ %MW1002 := %MW1305 ]  (* VSD1_CURRENT - par 0104 arus A x10 *)
  [ %MW1003 := %MW1308 ]  (* VSD1_DCBUS - par 0107 DC bus V *)
  [ %MW1004 := %MW1310 ]  (* VSD1_VOUT - par 0109 Vout V *)
  [ %MW1005 := %MW1312 ]  (* VSD1_REF_RB - par 0111 ext ref1 Hz x10 *)
  // as ST:
  //   VSD1_SW := %MW1302;
  //   VSD1_FREQ := %MW1304;
  //   VSD1_CURRENT := %MW1305;
  //   VSD1_DCBUS := %MW1308;
  //   VSD1_VOUT := %MW1310;
  //   VSD1_REF_RB := %MW1312;

// Rung 40: SCALE_VSD2
// VSD2 ACS580 -> FUXA. /40: 20000 = 46.02 = 50,00 Hz -> Hz x10
  LD 1
  [ %MW1020 := %MW1342 ]  (* VSD2_SW - status word *)
  [ %MW1021 := %MW1343 / 40 ](* VSD2_FREQ - act1 -> Hz x10 *)
  [ %MF1220 := DINT_TO_REAL( %MD1210 ) ](* 01.07 arus, 100 = 1 A *)
  [ %MF1220 := %MF1220 / 10.0 ]
  [ %MW1022 := REAL_TO_INT( %MF1220 ) ](* VSD2_CURRENT - arus A x10 *)
  [ %MW1023 := %MW1346 / 10 ](* VSD2_DCBUS - 01.11 DC bus V *)
  [ %MW1024 := %MW1347 ]  (* VSD2_VOUT - 01.13 Vout V *)
  [ %MW1025 := %MW1340 / 40 ](* VSD2_REF_RB - ref1 terbaca balik Hz x10 *)
  // as ST:
  //   VSD2_SW := %MW1342;
  //   VSD2_FREQ := %MW1343 / 40;
  //   %MF1220 := DINT_TO_REAL( %MD1210 );
  //   %MF1220 := %MF1220 / 10.0;
  //   VSD2_CURRENT := REAL_TO_INT( %MF1220 );
  //   VSD2_DCBUS := %MW1346 / 10;
  //   VSD2_VOUT := %MW1347;
  //   VSD2_REF_RB := %MW1340 / 40;

// Rung 41: SCALE_VSD3
// VSD3 ACS580 -> FUXA. /40: 20000 = 46.02 = 50,00 Hz -> Hz x10
  LD 1
  [ %MW1040 := %MW1382 ]  (* VSD3_SW - status word *)
  [ %MW1041 := %MW1383 / 40 ](* VSD3_FREQ - act1 -> Hz x10 *)
  [ %MF1222 := DINT_TO_REAL( %MD1212 ) ](* 01.07 arus, 100 = 1 A *)
  [ %MF1222 := %MF1222 / 10.0 ]
  [ %MW1042 := REAL_TO_INT( %MF1222 ) ](* VSD3_CURRENT - arus A x10 *)
  [ %MW1043 := %MW1386 / 10 ](* VSD3_DCBUS - 01.11 DC bus V *)
  [ %MW1044 := %MW1387 ]  (* VSD3_VOUT - 01.13 Vout V *)
  [ %MW1045 := %MW1380 / 40 ](* VSD3_REF_RB - ref1 terbaca balik Hz x10 *)
  // as ST:
  //   VSD3_SW := %MW1382;
  //   VSD3_FREQ := %MW1383 / 40;
  //   %MF1222 := DINT_TO_REAL( %MD1212 );
  //   %MF1222 := %MF1222 / 10.0;
  //   VSD3_CURRENT := REAL_TO_INT( %MF1222 );
  //   VSD3_DCBUS := %MW1386 / 10;
  //   VSD3_VOUT := %MW1387;
  //   VSD3_REF_RB := %MW1380 / 40;

// Rung 42: SCALE_VSD4
// VSD4 ACS580 -> FUXA. /40: 20000 = 46.02 = 50,00 Hz -> Hz x10
  LD 1
  [ %MW1060 := %MW1462 ]  (* VSD4_SW - status word *)
  [ %MW1061 := %MW1463 / 40 ](* VSD4_FREQ - act1 -> Hz x10 *)
  [ %MF1224 := DINT_TO_REAL( %MD1214 ) ](* 01.07 arus, 100 = 1 A *)
  [ %MF1224 := %MF1224 / 10.0 ]
  [ %MW1062 := REAL_TO_INT( %MF1224 ) ](* VSD4_CURRENT - arus A x10 *)
  [ %MW1063 := %MW1466 / 10 ](* VSD4_DCBUS - 01.11 DC bus V *)
  [ %MW1064 := %MW1467 ]  (* VSD4_VOUT - 01.13 Vout V *)
  [ %MW1065 := %MW1460 / 40 ](* VSD4_REF_RB - ref1 terbaca balik Hz x10 *)
  // as ST:
  //   VSD4_SW := %MW1462;
  //   VSD4_FREQ := %MW1463 / 40;
  //   %MF1224 := DINT_TO_REAL( %MD1214 );
  //   %MF1224 := %MF1224 / 10.0;
  //   VSD4_CURRENT := REAL_TO_INT( %MF1224 );
  //   VSD4_DCBUS := %MW1466 / 10;
  //   VSD4_VOUT := %MW1467;
  //   VSD4_REF_RB := %MW1460 / 40;

// Rung 43: SCALE_VSD5
// VSD5 ACS580 -> FUXA. /40: 20000 = 46.02 = 50,00 Hz -> Hz x10
  LD 1
  [ %MW1080 := %MW1502 ]  (* VSD5_SW - status word *)
  [ %MW1081 := %MW1503 / 40 ](* VSD5_FREQ - act1 -> Hz x10 *)
  [ %MF1226 := DINT_TO_REAL( %MD1216 ) ](* 01.07 arus, 100 = 1 A *)
  [ %MF1226 := %MF1226 / 10.0 ]
  [ %MW1082 := REAL_TO_INT( %MF1226 ) ](* VSD5_CURRENT - arus A x10 *)
  [ %MW1083 := %MW1506 / 10 ](* VSD5_DCBUS - 01.11 DC bus V *)
  [ %MW1084 := %MW1507 ]  (* VSD5_VOUT - 01.13 Vout V *)
  [ %MW1085 := %MW1500 / 40 ](* VSD5_REF_RB - ref1 terbaca balik Hz x10 *)
  // as ST:
  //   VSD5_SW := %MW1502;
  //   VSD5_FREQ := %MW1503 / 40;
  //   %MF1226 := DINT_TO_REAL( %MD1216 );
  //   %MF1226 := %MF1226 / 10.0;
  //   VSD5_CURRENT := REAL_TO_INT( %MF1226 );
  //   VSD5_DCBUS := %MW1506 / 10;
  //   VSD5_VOUT := %MW1507;
  //   VSD5_REF_RB := %MW1500 / 40;

// Rung 44: STAT_RUN_VSD1
// VSD1 berjalan (status word bit 2 RDY_REF)
  LD %MW1000:X2           (* VSD1_SW *)
  ST %M25                 (* VSD1_RUNNING *)
  // as ST:
  //   VSD1_RUNNING := VSD1_SW:X2;

// Rung 45: STAT_FLT_VSD1
// VSD1 FAULT (bit 3 TRIPPED), hanya dipercaya bila komunikasi OK
  LD %M60                 (* VSD1_COMM_OK - COMM_OK *)
  AND %MW1000:X3          (* VSD1_SW *)
  ST %M40                 (* VSD1_FAULT *)
  // as ST:
  //   VSD1_FAULT := VSD1_COMM_OK AND VSD1_SW:X3;

// Rung 46: STAT_WRN_VSD1
// VSD1 warning (bit 7 ALARM)
  LD %MW1000:X7           (* VSD1_SW *)
  ST %M45                 (* VSD1_WARN *)
  // as ST:
  //   VSD1_WARN := VSD1_SW:X7;

// Rung 47: STAT_REM_VSD1
// VSD1 di REMOTE (bit 9)
  LD %MW1000:X9           (* VSD1_SW *)
  ST %M50                 (* VSD1_REMOTE *)
  // as ST:
  //   VSD1_REMOTE := VSD1_SW:X9;

// Rung 48: STAT_RUN_VSD2
// VSD2 berjalan (status word bit 2 RDY_REF)
  LD %MW1020:X2           (* VSD2_SW *)
  ST %M26                 (* VSD2_RUNNING *)
  // as ST:
  //   VSD2_RUNNING := VSD2_SW:X2;

// Rung 49: STAT_FLT_VSD2
// VSD2 FAULT (bit 3 TRIPPED), hanya dipercaya bila komunikasi OK
  LD %M61                 (* VSD2_COMM_OK - COMM_OK *)
  AND %MW1020:X3          (* VSD2_SW *)
  ST %M41                 (* VSD2_FAULT *)
  // as ST:
  //   VSD2_FAULT := VSD2_COMM_OK AND VSD2_SW:X3;

// Rung 50: STAT_WRN_VSD2
// VSD2 warning (bit 7 ALARM)
  LD %MW1020:X7           (* VSD2_SW *)
  ST %M46                 (* VSD2_WARN *)
  // as ST:
  //   VSD2_WARN := VSD2_SW:X7;

// Rung 51: STAT_REM_VSD2
// VSD2 di REMOTE (bit 9)
  LD %MW1020:X9           (* VSD2_SW *)
  ST %M51                 (* VSD2_REMOTE *)
  // as ST:
  //   VSD2_REMOTE := VSD2_SW:X9;

// Rung 52: STAT_RUN_VSD3
// VSD3 berjalan (status word bit 2 RDY_REF)
  LD %MW1040:X2           (* VSD3_SW *)
  ST %M27                 (* VSD3_RUNNING *)
  // as ST:
  //   VSD3_RUNNING := VSD3_SW:X2;

// Rung 53: STAT_FLT_VSD3
// VSD3 FAULT (bit 3 TRIPPED), hanya dipercaya bila komunikasi OK
  LD %M62                 (* VSD3_COMM_OK - COMM_OK *)
  AND %MW1040:X3          (* VSD3_SW *)
  ST %M42                 (* VSD3_FAULT *)
  // as ST:
  //   VSD3_FAULT := VSD3_COMM_OK AND VSD3_SW:X3;

// Rung 54: STAT_WRN_VSD3
// VSD3 warning (bit 7 ALARM)
  LD %MW1040:X7           (* VSD3_SW *)
  ST %M47                 (* VSD3_WARN *)
  // as ST:
  //   VSD3_WARN := VSD3_SW:X7;

// Rung 55: STAT_REM_VSD3
// VSD3 di REMOTE (bit 9)
  LD %MW1040:X9           (* VSD3_SW *)
  ST %M52                 (* VSD3_REMOTE *)
  // as ST:
  //   VSD3_REMOTE := VSD3_SW:X9;

// Rung 56: STAT_RUN_VSD4
// VSD4 berjalan (status word bit 2 RDY_REF)
  LD %MW1060:X2           (* VSD4_SW *)
  ST %M28                 (* VSD4_RUNNING *)
  // as ST:
  //   VSD4_RUNNING := VSD4_SW:X2;

// Rung 57: STAT_FLT_VSD4
// VSD4 FAULT (bit 3 TRIPPED), hanya dipercaya bila komunikasi OK
  LD %M63                 (* VSD4_COMM_OK - COMM_OK *)
  AND %MW1060:X3          (* VSD4_SW *)
  ST %M43                 (* VSD4_FAULT *)
  // as ST:
  //   VSD4_FAULT := VSD4_COMM_OK AND VSD4_SW:X3;

// Rung 58: STAT_WRN_VSD4
// VSD4 warning (bit 7 ALARM)
  LD %MW1060:X7           (* VSD4_SW *)
  ST %M48                 (* VSD4_WARN *)
  // as ST:
  //   VSD4_WARN := VSD4_SW:X7;

// Rung 59: STAT_REM_VSD4
// VSD4 di REMOTE (bit 9)
  LD %MW1060:X9           (* VSD4_SW *)
  ST %M53                 (* VSD4_REMOTE *)
  // as ST:
  //   VSD4_REMOTE := VSD4_SW:X9;

// Rung 60: STAT_RUN_VSD5
// VSD5 berjalan (status word bit 2 RDY_REF)
  LD %MW1080:X2           (* VSD5_SW *)
  ST %M29                 (* VSD5_RUNNING *)
  // as ST:
  //   VSD5_RUNNING := VSD5_SW:X2;

// Rung 61: STAT_FLT_VSD5
// VSD5 FAULT (bit 3 TRIPPED), hanya dipercaya bila komunikasi OK
  LD %M64                 (* VSD5_COMM_OK - COMM_OK *)
  AND %MW1080:X3          (* VSD5_SW *)
  ST %M44                 (* VSD5_FAULT *)
  // as ST:
  //   VSD5_FAULT := VSD5_COMM_OK AND VSD5_SW:X3;

// Rung 62: STAT_WRN_VSD5
// VSD5 warning (bit 7 ALARM)
  LD %MW1080:X7           (* VSD5_SW *)
  ST %M49                 (* VSD5_WARN *)
  // as ST:
  //   VSD5_WARN := VSD5_SW:X7;

// Rung 63: STAT_REM_VSD5
// VSD5 di REMOTE (bit 9)
  LD %MW1080:X9           (* VSD5_SW *)
  ST %M54                 (* VSD5_REMOTE *)
  // as ST:
  //   VSD5_REMOTE := VSD5_SW:X9;

// Rung 64: SP_MAX_VSD1
// VSD1 setpoint dari FUXA (%MW1006, Hz x10) dibatasi SP_MAX
  LD [ %MW1006 > %MW991 ] (* VSD1_SP, SP_MAX *)
  [ %MW1006 := %MW991 ]   (* VSD1_SP, SP_MAX *)
  // as ST:
  //   IF VSD1_SP > SP_MAX THEN VSD1_SP := SP_MAX; END_IF;

// Rung 65: SP_MIN_VSD1
// VSD1 setpoint dibatasi SP_MIN
  LD [ %MW1006 < %MW990 ] (* VSD1_SP, SP_MIN *)
  [ %MW1006 := %MW990 ]   (* VSD1_SP, SP_MIN *)
  // as ST:
  //   IF VSD1_SP < SP_MIN THEN VSD1_SP := SP_MIN; END_IF;

// Rung 66: SP_REF_VSD1
// VSD1 ref1 ke drive: Hz x10 * 40 (20000 = 50 Hz). Ditulis IOScanner tiap 500 ms
  LD 1
  [ %MW1251 := %MW1006 * 40 ](* VSD1_SP *)
  [ %QWN100.2.0 := %MW1251 ]
  // as ST:
  //   %MW1251 := VSD1_SP * 40;
  //   %QWN100.2.0 := %MW1251;

// Rung 67: SP_MAX_VSD2
// VSD2 setpoint dari FUXA (%MW1026, Hz x10) dibatasi SP_MAX
  LD [ %MW1026 > %MW991 ] (* VSD2_SP, SP_MAX *)
  [ %MW1026 := %MW991 ]   (* VSD2_SP, SP_MAX *)
  // as ST:
  //   IF VSD2_SP > SP_MAX THEN VSD2_SP := SP_MAX; END_IF;

// Rung 68: SP_MIN_VSD2
// VSD2 setpoint dibatasi SP_MIN
  LD [ %MW1026 < %MW990 ] (* VSD2_SP, SP_MIN *)
  [ %MW1026 := %MW990 ]   (* VSD2_SP, SP_MIN *)
  // as ST:
  //   IF VSD2_SP < SP_MIN THEN VSD2_SP := SP_MIN; END_IF;

// Rung 69: SP_REF_VSD2
// VSD2 ref1 ke drive: Hz x10 * 40 (20000 = 50 Hz). Ditulis IOScanner tiap 500 ms
  LD 1
  [ %MW1252 := %MW1026 * 40 ](* VSD2_SP *)
  [ %QWN101.4.0 := %MW1252 ]
  // as ST:
  //   %MW1252 := VSD2_SP * 40;
  //   %QWN101.4.0 := %MW1252;

// Rung 70: SP_MAX_VSD3
// VSD3 setpoint dari FUXA (%MW1046, Hz x10) dibatasi SP_MAX
  LD [ %MW1046 > %MW991 ] (* VSD3_SP, SP_MAX *)
  [ %MW1046 := %MW991 ]   (* VSD3_SP, SP_MAX *)
  // as ST:
  //   IF VSD3_SP > SP_MAX THEN VSD3_SP := SP_MAX; END_IF;

// Rung 71: SP_MIN_VSD3
// VSD3 setpoint dibatasi SP_MIN
  LD [ %MW1046 < %MW990 ] (* VSD3_SP, SP_MIN *)
  [ %MW1046 := %MW990 ]   (* VSD3_SP, SP_MIN *)
  // as ST:
  //   IF VSD3_SP < SP_MIN THEN VSD3_SP := SP_MIN; END_IF;

// Rung 72: SP_REF_VSD3
// VSD3 ref1 ke drive: Hz x10 * 40 (20000 = 50 Hz). Ditulis IOScanner tiap 500 ms
  LD 1
  [ %MW1253 := %MW1046 * 40 ](* VSD3_SP *)
  [ %QWN102.4.0 := %MW1253 ]
  // as ST:
  //   %MW1253 := VSD3_SP * 40;
  //   %QWN102.4.0 := %MW1253;

// Rung 73: SP_MAX_VSD4
// VSD4 setpoint dari FUXA (%MW1066, Hz x10) dibatasi SP_MAX
  LD [ %MW1066 > %MW991 ] (* VSD4_SP, SP_MAX *)
  [ %MW1066 := %MW991 ]   (* VSD4_SP, SP_MAX *)
  // as ST:
  //   IF VSD4_SP > SP_MAX THEN VSD4_SP := SP_MAX; END_IF;

// Rung 74: SP_MIN_VSD4
// VSD4 setpoint dibatasi SP_MIN
  LD [ %MW1066 < %MW990 ] (* VSD4_SP, SP_MIN *)
  [ %MW1066 := %MW990 ]   (* VSD4_SP, SP_MIN *)
  // as ST:
  //   IF VSD4_SP < SP_MIN THEN VSD4_SP := SP_MIN; END_IF;

// Rung 75: SP_REF_VSD4
// VSD4 ref1 ke drive: Hz x10 * 40 (20000 = 50 Hz). Ditulis IOScanner tiap 500 ms
  LD 1
  [ %MW1254 := %MW1066 * 40 ](* VSD4_SP *)
  [ %QWN104.4.0 := %MW1254 ]
  // as ST:
  //   %MW1254 := VSD4_SP * 40;
  //   %QWN104.4.0 := %MW1254;

// Rung 76: SP_MAX_VSD5
// VSD5 setpoint dari FUXA (%MW1086, Hz x10) dibatasi SP_MAX
  LD [ %MW1086 > %MW991 ] (* VSD5_SP, SP_MAX *)
  [ %MW1086 := %MW991 ]   (* VSD5_SP, SP_MAX *)
  // as ST:
  //   IF VSD5_SP > SP_MAX THEN VSD5_SP := SP_MAX; END_IF;

// Rung 77: SP_MIN_VSD5
// VSD5 setpoint dibatasi SP_MIN
  LD [ %MW1086 < %MW990 ] (* VSD5_SP, SP_MIN *)
  [ %MW1086 := %MW990 ]   (* VSD5_SP, SP_MIN *)
  // as ST:
  //   IF VSD5_SP < SP_MIN THEN VSD5_SP := SP_MIN; END_IF;

// Rung 78: SP_REF_VSD5
// VSD5 ref1 ke drive: Hz x10 * 40 (20000 = 50 Hz). Ditulis IOScanner tiap 500 ms
  LD 1
  [ %MW1255 := %MW1086 * 40 ](* VSD5_SP *)
  [ %QWN105.4.0 := %MW1255 ]
  // as ST:
  //   %MW1255 := VSD5_SP * 40;
  //   %QWN105.4.0 := %MW1255;

// Rung 79: START_REM_VSD1
// VSD1 START dari SCADA (%M10): hanya di REMOTE, ditolak bila fault / PB OFF ditekan
  LD %I0.0                (* SEL_REMOTE - REMOTE *)
  AND %M10                (* VSD1_START - START FUXA *)
  AND %I0.3               (* VSD1_PB_OFF - PB OFF tidak ditekan (NC) *)
  ANDN %M40               (* VSD1_FAULT - tidak fault *)
  S %Q0.0                 (* VSD1_RUN *)
  // as ST:
  //   IF SEL_REMOTE AND VSD1_START AND VSD1_PB_OFF AND NOT VSD1_FAULT THEN VSD1_RUN := TRUE; END_IF;

// Rung 80: START_LOC_VSD1
// VSD1 START dari PB ON panel (%I0.2): hanya di LOCAL, ditolak bila fault / PB OFF ditekan
  LDN %I0.0               (* SEL_REMOTE - LOCAL *)
  AND %I0.2               (* VSD1_PB_ON - PB ON (NO) *)
  AND %I0.3               (* VSD1_PB_OFF - PB OFF tidak ditekan (NC) *)
  ANDN %M40               (* VSD1_FAULT - tidak fault *)
  S %Q0.0                 (* VSD1_RUN *)
  // as ST:
  //   IF NOT SEL_REMOTE AND VSD1_PB_ON AND VSD1_PB_OFF AND NOT VSD1_FAULT THEN VSD1_RUN := TRUE; END_IF;

// Rung 81: STOP_REM_VSD1
// VSD1 STOP dari SCADA (%M11): hanya di REMOTE
  LD %I0.0                (* SEL_REMOTE - REMOTE *)
  AND %M11                (* VSD1_STOP - STOP FUXA *)
  R %Q0.0                 (* VSD1_RUN *)
  // as ST:
  //   IF SEL_REMOTE AND VSD1_STOP THEN VSD1_RUN := FALSE; END_IF;

// Rung 82: STOP_PB_VSD1
// VSD1 STOP dari PB OFF panel (%I0.3, NC): aktif di LOCAL dan REMOTE; kabel putus = stop
  LDN %I0.3               (* VSD1_PB_OFF - PB OFF ditekan / kabel putus *)
  R %Q0.0                 (* VSD1_RUN *)
  // as ST:
  //   IF NOT VSD1_PB_OFF THEN VSD1_RUN := FALSE; END_IF;

// Rung 83: STOP_FLT_VSD1
// VSD1 fault (status word, comm OK) -> RUN mati
  LD %M40                 (* VSD1_FAULT *)
  R %Q0.0                 (* VSD1_RUN *)
  // as ST:
  //   IF VSD1_FAULT THEN VSD1_RUN := FALSE; END_IF;

// Rung 84: CLR_START_VSD1
// VSD1 bersihkan bit START dari FUXA (pulse; juga di LOCAL supaya tidak tertahan)
  LD %M10                 (* VSD1_START *)
  R %M10                  (* VSD1_START *)
  // as ST:
  //   IF VSD1_START THEN VSD1_START := FALSE; END_IF;

// Rung 85: CLR_STOP_VSD1
// VSD1 bersihkan bit STOP dari FUXA (pulse)
  LD %M11                 (* VSD1_STOP *)
  R %M11                  (* VSD1_STOP *)
  // as ST:
  //   IF VSD1_STOP THEN VSD1_STOP := FALSE; END_IF;

// Rung 86: START_REM_VSD2
// VSD2 START dari SCADA (%M12): hanya di REMOTE, ditolak bila fault / PB OFF ditekan
  LD %I0.0                (* SEL_REMOTE - REMOTE *)
  AND %M12                (* VSD2_START - START FUXA *)
  AND %I0.5               (* VSD2_PB_OFF - PB OFF tidak ditekan (NC) *)
  ANDN %M41               (* VSD2_FAULT - tidak fault *)
  S %Q0.1                 (* VSD2_RUN *)
  // as ST:
  //   IF SEL_REMOTE AND VSD2_START AND VSD2_PB_OFF AND NOT VSD2_FAULT THEN VSD2_RUN := TRUE; END_IF;

// Rung 87: START_LOC_VSD2
// VSD2 START dari PB ON panel (%I0.4): hanya di LOCAL, ditolak bila fault / PB OFF ditekan
  LDN %I0.0               (* SEL_REMOTE - LOCAL *)
  AND %I0.4               (* VSD2_PB_ON - PB ON (NO) *)
  AND %I0.5               (* VSD2_PB_OFF - PB OFF tidak ditekan (NC) *)
  ANDN %M41               (* VSD2_FAULT - tidak fault *)
  S %Q0.1                 (* VSD2_RUN *)
  // as ST:
  //   IF NOT SEL_REMOTE AND VSD2_PB_ON AND VSD2_PB_OFF AND NOT VSD2_FAULT THEN VSD2_RUN := TRUE; END_IF;

// Rung 88: STOP_REM_VSD2
// VSD2 STOP dari SCADA (%M13): hanya di REMOTE
  LD %I0.0                (* SEL_REMOTE - REMOTE *)
  AND %M13                (* VSD2_STOP - STOP FUXA *)
  R %Q0.1                 (* VSD2_RUN *)
  // as ST:
  //   IF SEL_REMOTE AND VSD2_STOP THEN VSD2_RUN := FALSE; END_IF;

// Rung 89: STOP_PB_VSD2
// VSD2 STOP dari PB OFF panel (%I0.5, NC): aktif di LOCAL dan REMOTE; kabel putus = stop
  LDN %I0.5               (* VSD2_PB_OFF - PB OFF ditekan / kabel putus *)
  R %Q0.1                 (* VSD2_RUN *)
  // as ST:
  //   IF NOT VSD2_PB_OFF THEN VSD2_RUN := FALSE; END_IF;

// Rung 90: STOP_FLT_VSD2
// VSD2 fault (status word, comm OK) -> RUN mati
  LD %M41                 (* VSD2_FAULT *)
  R %Q0.1                 (* VSD2_RUN *)
  // as ST:
  //   IF VSD2_FAULT THEN VSD2_RUN := FALSE; END_IF;

// Rung 91: CLR_START_VSD2
// VSD2 bersihkan bit START dari FUXA (pulse; juga di LOCAL supaya tidak tertahan)
  LD %M12                 (* VSD2_START *)
  R %M12                  (* VSD2_START *)
  // as ST:
  //   IF VSD2_START THEN VSD2_START := FALSE; END_IF;

// Rung 92: CLR_STOP_VSD2
// VSD2 bersihkan bit STOP dari FUXA (pulse)
  LD %M13                 (* VSD2_STOP *)
  R %M13                  (* VSD2_STOP *)
  // as ST:
  //   IF VSD2_STOP THEN VSD2_STOP := FALSE; END_IF;

// Rung 93: START_REM_VSD3
// VSD3 START dari SCADA (%M14): hanya di REMOTE, ditolak bila fault / PB OFF ditekan
  LD %I0.0                (* SEL_REMOTE - REMOTE *)
  AND %M14                (* VSD3_START - START FUXA *)
  AND %I0.7               (* VSD3_PB_OFF - PB OFF tidak ditekan (NC) *)
  ANDN %M42               (* VSD3_FAULT - tidak fault *)
  S %Q0.2                 (* VSD3_RUN *)
  // as ST:
  //   IF SEL_REMOTE AND VSD3_START AND VSD3_PB_OFF AND NOT VSD3_FAULT THEN VSD3_RUN := TRUE; END_IF;

// Rung 94: START_LOC_VSD3
// VSD3 START dari PB ON panel (%I0.6): hanya di LOCAL, ditolak bila fault / PB OFF ditekan
  LDN %I0.0               (* SEL_REMOTE - LOCAL *)
  AND %I0.6               (* VSD3_PB_ON - PB ON (NO) *)
  AND %I0.7               (* VSD3_PB_OFF - PB OFF tidak ditekan (NC) *)
  ANDN %M42               (* VSD3_FAULT - tidak fault *)
  S %Q0.2                 (* VSD3_RUN *)
  // as ST:
  //   IF NOT SEL_REMOTE AND VSD3_PB_ON AND VSD3_PB_OFF AND NOT VSD3_FAULT THEN VSD3_RUN := TRUE; END_IF;

// Rung 95: STOP_REM_VSD3
// VSD3 STOP dari SCADA (%M15): hanya di REMOTE
  LD %I0.0                (* SEL_REMOTE - REMOTE *)
  AND %M15                (* VSD3_STOP - STOP FUXA *)
  R %Q0.2                 (* VSD3_RUN *)
  // as ST:
  //   IF SEL_REMOTE AND VSD3_STOP THEN VSD3_RUN := FALSE; END_IF;

// Rung 96: STOP_PB_VSD3
// VSD3 STOP dari PB OFF panel (%I0.7, NC): aktif di LOCAL dan REMOTE; kabel putus = stop
  LDN %I0.7               (* VSD3_PB_OFF - PB OFF ditekan / kabel putus *)
  R %Q0.2                 (* VSD3_RUN *)
  // as ST:
  //   IF NOT VSD3_PB_OFF THEN VSD3_RUN := FALSE; END_IF;

// Rung 97: STOP_FLT_VSD3
// VSD3 fault (status word, comm OK) -> RUN mati
  LD %M42                 (* VSD3_FAULT *)
  R %Q0.2                 (* VSD3_RUN *)
  // as ST:
  //   IF VSD3_FAULT THEN VSD3_RUN := FALSE; END_IF;

// Rung 98: CLR_START_VSD3
// VSD3 bersihkan bit START dari FUXA (pulse; juga di LOCAL supaya tidak tertahan)
  LD %M14                 (* VSD3_START *)
  R %M14                  (* VSD3_START *)
  // as ST:
  //   IF VSD3_START THEN VSD3_START := FALSE; END_IF;

// Rung 99: CLR_STOP_VSD3
// VSD3 bersihkan bit STOP dari FUXA (pulse)
  LD %M15                 (* VSD3_STOP *)
  R %M15                  (* VSD3_STOP *)
  // as ST:
  //   IF VSD3_STOP THEN VSD3_STOP := FALSE; END_IF;

// Rung 100: START_REM_VSD4
// VSD4 START dari SCADA (%M16): hanya di REMOTE, ditolak bila fault / PB OFF ditekan
  LD %I0.0                (* SEL_REMOTE - REMOTE *)
  AND %M16                (* VSD4_START - START FUXA *)
  AND %I0.9               (* VSD4_PB_OFF - PB OFF tidak ditekan (NC) *)
  ANDN %M43               (* VSD4_FAULT - tidak fault *)
  S %Q0.3                 (* VSD4_RUN *)
  // as ST:
  //   IF SEL_REMOTE AND VSD4_START AND VSD4_PB_OFF AND NOT VSD4_FAULT THEN VSD4_RUN := TRUE; END_IF;

// Rung 101: START_LOC_VSD4
// VSD4 START dari PB ON panel (%I0.8): hanya di LOCAL, ditolak bila fault / PB OFF ditekan
  LDN %I0.0               (* SEL_REMOTE - LOCAL *)
  AND %I0.8               (* VSD4_PB_ON - PB ON (NO) *)
  AND %I0.9               (* VSD4_PB_OFF - PB OFF tidak ditekan (NC) *)
  ANDN %M43               (* VSD4_FAULT - tidak fault *)
  S %Q0.3                 (* VSD4_RUN *)
  // as ST:
  //   IF NOT SEL_REMOTE AND VSD4_PB_ON AND VSD4_PB_OFF AND NOT VSD4_FAULT THEN VSD4_RUN := TRUE; END_IF;

// Rung 102: STOP_REM_VSD4
// VSD4 STOP dari SCADA (%M17): hanya di REMOTE
  LD %I0.0                (* SEL_REMOTE - REMOTE *)
  AND %M17                (* VSD4_STOP - STOP FUXA *)
  R %Q0.3                 (* VSD4_RUN *)
  // as ST:
  //   IF SEL_REMOTE AND VSD4_STOP THEN VSD4_RUN := FALSE; END_IF;

// Rung 103: STOP_PB_VSD4
// VSD4 STOP dari PB OFF panel (%I0.9, NC): aktif di LOCAL dan REMOTE; kabel putus = stop
  LDN %I0.9               (* VSD4_PB_OFF - PB OFF ditekan / kabel putus *)
  R %Q0.3                 (* VSD4_RUN *)
  // as ST:
  //   IF NOT VSD4_PB_OFF THEN VSD4_RUN := FALSE; END_IF;

// Rung 104: STOP_FLT_VSD4
// VSD4 fault (status word, comm OK) -> RUN mati
  LD %M43                 (* VSD4_FAULT *)
  R %Q0.3                 (* VSD4_RUN *)
  // as ST:
  //   IF VSD4_FAULT THEN VSD4_RUN := FALSE; END_IF;

// Rung 105: CLR_START_VSD4
// VSD4 bersihkan bit START dari FUXA (pulse; juga di LOCAL supaya tidak tertahan)
  LD %M16                 (* VSD4_START *)
  R %M16                  (* VSD4_START *)
  // as ST:
  //   IF VSD4_START THEN VSD4_START := FALSE; END_IF;

// Rung 106: CLR_STOP_VSD4
// VSD4 bersihkan bit STOP dari FUXA (pulse)
  LD %M17                 (* VSD4_STOP *)
  R %M17                  (* VSD4_STOP *)
  // as ST:
  //   IF VSD4_STOP THEN VSD4_STOP := FALSE; END_IF;

// Rung 107: START_REM_VSD5
// VSD5 START dari SCADA (%M18): hanya di REMOTE, ditolak bila fault / PB OFF ditekan
  LD %I0.0                (* SEL_REMOTE - REMOTE *)
  AND %M18                (* VSD5_START - START FUXA *)
  AND %I0.11              (* VSD5_PB_OFF - PB OFF tidak ditekan (NC) *)
  ANDN %M44               (* VSD5_FAULT - tidak fault *)
  S %Q0.4                 (* VSD5_RUN *)
  // as ST:
  //   IF SEL_REMOTE AND VSD5_START AND VSD5_PB_OFF AND NOT VSD5_FAULT THEN VSD5_RUN := TRUE; END_IF;

// Rung 108: START_LOC_VSD5
// VSD5 START dari PB ON panel (%I0.10): hanya di LOCAL, ditolak bila fault / PB OFF ditekan
  LDN %I0.0               (* SEL_REMOTE - LOCAL *)
  AND %I0.10              (* VSD5_PB_ON - PB ON (NO) *)
  AND %I0.11              (* VSD5_PB_OFF - PB OFF tidak ditekan (NC) *)
  ANDN %M44               (* VSD5_FAULT - tidak fault *)
  S %Q0.4                 (* VSD5_RUN *)
  // as ST:
  //   IF NOT SEL_REMOTE AND VSD5_PB_ON AND VSD5_PB_OFF AND NOT VSD5_FAULT THEN VSD5_RUN := TRUE; END_IF;

// Rung 109: STOP_REM_VSD5
// VSD5 STOP dari SCADA (%M19): hanya di REMOTE
  LD %I0.0                (* SEL_REMOTE - REMOTE *)
  AND %M19                (* VSD5_STOP - STOP FUXA *)
  R %Q0.4                 (* VSD5_RUN *)
  // as ST:
  //   IF SEL_REMOTE AND VSD5_STOP THEN VSD5_RUN := FALSE; END_IF;

// Rung 110: STOP_PB_VSD5
// VSD5 STOP dari PB OFF panel (%I0.11, NC): aktif di LOCAL dan REMOTE; kabel putus = stop
  LDN %I0.11              (* VSD5_PB_OFF - PB OFF ditekan / kabel putus *)
  R %Q0.4                 (* VSD5_RUN *)
  // as ST:
  //   IF NOT VSD5_PB_OFF THEN VSD5_RUN := FALSE; END_IF;

// Rung 111: STOP_FLT_VSD5
// VSD5 fault (status word, comm OK) -> RUN mati
  LD %M44                 (* VSD5_FAULT *)
  R %Q0.4                 (* VSD5_RUN *)
  // as ST:
  //   IF VSD5_FAULT THEN VSD5_RUN := FALSE; END_IF;

// Rung 112: CLR_START_VSD5
// VSD5 bersihkan bit START dari FUXA (pulse; juga di LOCAL supaya tidak tertahan)
  LD %M18                 (* VSD5_START *)
  R %M18                  (* VSD5_START *)
  // as ST:
  //   IF VSD5_START THEN VSD5_START := FALSE; END_IF;

// Rung 113: CLR_STOP_VSD5
// VSD5 bersihkan bit STOP dari FUXA (pulse)
  LD %M19                 (* VSD5_STOP *)
  R %M19                  (* VSD5_STOP *)
  // as ST:
  //   IF VSD5_STOP THEN VSD5_STOP := FALSE; END_IF;

// Rung 114: INTERLOCK
// E-stop tidak sehat (%I0.1 = 0) -> semua RUN mati. Selector TIDAK lagi menghentikan pompa (bumpless). HARUS di bawah rung START
  LDN %I0.1               (* ESTOP_OK - ESTOP_OK (NC) *)
  R %Q0.0                 (* VSD1_RUN *)
  R %Q0.1                 (* VSD2_RUN *)
  R %Q0.2                 (* VSD3_RUN *)
  R %Q0.3                 (* VSD4_RUN *)
  R %Q0.4                 (* VSD5_RUN *)
  // as ST:
  //   IF NOT ESTOP_OK THEN VSD1_RUN := FALSE; END_IF;
  //   IF NOT ESTOP_OK THEN VSD2_RUN := FALSE; END_IF;
  //   IF NOT ESTOP_OK THEN VSD3_RUN := FALSE; END_IF;
  //   IF NOT ESTOP_OK THEN VSD4_RUN := FALSE; END_IF;
  //   IF NOT ESTOP_OK THEN VSD5_RUN := FALSE; END_IF;

// Rung 115: MODE_REMOTE
// Status selector untuk FUXA: %M30 = 1 REMOTE, 0 LOCAL (FUXA menonaktifkan tombol START/STOP saat LOCAL)
  LD %I0.0                (* SEL_REMOTE *)
  ST %M30                 (* MODE_REMOTE *)
  // as ST:
  //   MODE_REMOTE := SEL_REMOTE;

// Rung 116: MODE_ESTOP
// Status e-stop untuk FUXA: %M31 = 1 sehat
  LD %I0.1                (* ESTOP_OK *)
  ST %M31                 (* MODE_ESTOP_OK *)
  // as ST:
  //   MODE_ESTOP_OK := ESTOP_OK;

// Rung 117: RUN_FB_VSD1
// Umpan balik output RUN VSD1 untuk FUXA
  LD %Q0.0                (* VSD1_RUN *)
  ST %M20                 (* VSD1_RUN_CMD *)
  // as ST:
  //   VSD1_RUN_CMD := VSD1_RUN;

// Rung 118: RUN_FB_VSD2
// Umpan balik output RUN VSD2 untuk FUXA
  LD %Q0.1                (* VSD2_RUN *)
  ST %M21                 (* VSD2_RUN_CMD *)
  // as ST:
  //   VSD2_RUN_CMD := VSD2_RUN;

// Rung 119: RUN_FB_VSD3
// Umpan balik output RUN VSD3 untuk FUXA
  LD %Q0.2                (* VSD3_RUN *)
  ST %M22                 (* VSD3_RUN_CMD *)
  // as ST:
  //   VSD3_RUN_CMD := VSD3_RUN;

// Rung 120: RUN_FB_VSD4
// Umpan balik output RUN VSD4 untuk FUXA
  LD %Q0.3                (* VSD4_RUN *)
  ST %M23                 (* VSD4_RUN_CMD *)
  // as ST:
  //   VSD4_RUN_CMD := VSD4_RUN;

// Rung 121: RUN_FB_VSD5
// Umpan balik output RUN VSD5 untuk FUXA
  LD %Q0.4                (* VSD5_RUN *)
  ST %M24                 (* VSD5_RUN_CMD *)
  // as ST:
  //   VSD5_RUN_CMD := VSD5_RUN;
